# EPICS substitutions: iocs/motor/acstech80-ioc/db/SPiiPlus.substitutions
# C's iocAcsTech80 SPiiPlus.substitutions, P and C from st.cmd.
file "$(MOTOR)/db/motor.db"
{
pattern
{N, M,       DTYP,       S, DESC,          EGU, DIR, VELO, VBAS, ACCL, BDST, BVEL, BACC, MRES, PREC, DHLM, DLLM, INIT}
{1, "m$(N)", "SPiiPlus", 0, "Motor M$(N)", mm,  Pos, 10,   0.,   1.,   0,    1,    .2,   1e-3, 3,    100,  -100, ""}
{2, "m$(N)", "SPiiPlus", 1, "Motor M$(N)", mm,  Pos, 10,   0.,   1.,   0,    1,    .2,   1e-3, 3,    100,  -100, ""}
}
